Fanuc KAREL source: KA00088.KL

PROGRAM KA00088
%NOLOCKGROUP
VAR
  SRC: JOINTPOS
  DST: STRING[80]
BEGIN
  DST = SRC
END KA00088
